Fanuc KAREL source: KT00250.KL

PROGRAM KT00250
%NOLOCKGROUP
VAR
  H1: ARRAY[2] OF SHORT
  B2: BOOLEAN
  OUT: INTEGER
BEGIN
  H1[1] = 2
    B2 = FALSE
  OUT = H1[1] OR B2
END KT00250
